PROGRAM MAIN
VAR
	Switch AT %I* :BOOL;
	LIGHT AT %Q* : BOOL;
END_VAR

Light := Switch;

END_PROGRAM

(* stored: Version 1.1.0.1
   POU MAIN: Id {f5350466-b198-4d8c-9e40-5bb2dc1b6287}, SpecialFunc None *)
